// TIA Portal V21 export
// export: Created 2026-11-10T19:39:05.8156129Z, ExportSetting WithDefaults, DisplayName Totally Integrated Automation Portal, DisplayVersion V21 Update 3, DisplayName STEP 7 Professional, DisplayVersion V21 Update 3, DisplayName STEP 7 Safety, DisplayVersion V21, DisplayName Tech WebApplication, DisplayVersion V21, DisplayName WinCC Basic/Comfort/Advanced, DisplayVersion V21 Update 3, DisplayName WinCC Unified, DisplayVersion V21 Update 3
DATA_BLOCK "DB_Common"   // DB1
{ S7_Optimized_Access := 'TRUE' }
VERSION : 0.1
// stored: AutoNumber true, DBAccessibleFromOPCUA true, DBAccessibleFromWebserver true, IsOnlyStoredInLoadMemory false, IsRetainMemResEnabled false, IsWriteProtectedInAS false, MemoryReserve 100
   VAR
      a_onlyA : Int;
      speed : Real := 1.5;
      flags : Array[0..7] of Bool;
      cfg : Struct
         ip : Array[0..3] of Byte;
         "name" : String[20] := 'PLC_A';
      END_STRUCT;
   END_VAR
BEGIN
END_DATA_BLOCK
